(* IEC 61131-3 sources: Lasal-MCP/examples/SampleSource/LASALScreenAdvancedSolution/LASALScreenAdvancedSolution/LASALScreenAdvacnedSolution/Stations/Terminal/HMI/Class/IconDestList, 1 file *)

(* ---- IconDestList.st ---- *)
(*!
<Class
	Name               = "IconDestList"
	Revision           = "0.0"
	RealtimeTask       = "false"
	CyclicTask         = "false"
	BackgroundTask     = "false"
	Sigmatek           = "false"
	OSInterface        = "false"
	HighPriority       = "false"
	Automatic          = "false"
	UpdateMode         = "Prescan"
	SharedCommandTable = "true"
	Objectsize         = "(540,420)">
	<Channels>
		<Client Name="_Grafix" Required="false" Internal="false"/>
		<Client Name="DragDropArea" Required="true" Internal="false"/>
		<Client Name="SigCLib" Required="false" Internal="false"/>
	</Channels>
	<Network Name="IconDestList">
		<!-- List of Components in this network -->
		<Components>
			<Object
				Name       = "_base"
				Class      = "_ScrollArea2"
				Position   = "(218,120)"
				Visualized = "true"
				Remotely   = "true">
				<Channels>
					<Server Name="ActPos"/>
					<Server Name="Refresh"/>
					<Server Name="Server0"/>
					<Client Name="ExtendedScrollBar" Value="0"/>
					<Client Name="LineHighness"/>
					<Client Name="LineWidth"/>
					<Client Name="Lse"/>
					<Client Name="VerticalLevel"/>
				</Channels>
			</Object>
		</Components>
		<Comments>
		</Comments>
		<!-- List of Connections in this network -->
		<Connections>
			<Connection Source="this.Server0" Destination="_base.Server0" Vertices="(886,210),(714,210),"/>
			<Connection Source="this.Refresh" Destination="_base.Refresh" Vertices="(886,270),(714,270),"/>
			<Connection Source="this.ActPos" Destination="_base.ActPos" Vertices="(886,330),(714,330),"/>
			<Connection Source="_base.Lse" Destination="this.Lse" Vertices="(218,210),(38,210),"/>
			<Connection Source="_base.VerticalLevel" Destination="this.VerticalLevel" Vertices="(218,270),(38,270),"/>
			<Connection Source="_base.LineWidth" Destination="this.LineWidth" Vertices="(218,330),(38,330),"/>
		</Connections>
		<!-- Headerfiles -->
		<Options>
		</Options>
	</Network>
</Class>
*)
#pragma using _ScrollArea2

IconDestList : CLASS
: _ScrollArea2
  //Servers:
  //Clients:
	DragDropArea 	: CltChCmd_DragDropArea;
	_Grafix 	: CltChCmd__Grafix;
	SigCLib 	: CltChCmd_SigCLib;
  //Variables:
		TextColor 	: _COLOR;
		FrameColor 	: _COLOR;
		BackgroundColor 	: _COLOR;
		myPioScroll 	: _SCROLL;
		myImageRoom 	: _ROOM;
		Lines : ARRAY [0..100] OF DINT;

		pLSEpio 	: ^_IO;
  //Functions:

	FUNCTION VIRTUAL GLOBAL Init;
				//! <Function Comment="[#ENGLISH]&#13;&#10;method is called cyclic during object is on screen&#13;&#10;&#13;&#10;pio ....... pointer to io information&#13;&#10;input .... TRUE it&apos;s an input / FALSE it&apos;s an output&#13;&#10;" Name="IF_Run"/>
	FUNCTION __CDECL VIRTUAL GLOBAL IF_Run
		VAR_INPUT
			pio 	: ^_IO;			//! <Variable Comment="pointer to _IO information given by LSE" Name="IF_Run.pio"/>
			input 	: BOOL;			//! <Variable Comment="TRUE it&apos;s an input&#13;&#10;FALSE it&apos;s an output" Name="IF_Run.input"/>
		END_VAR;
				//! <Function Comment="method is called every time when redraw of a single line is necessary.&#13;&#10;" Name="Line"/>
	FUNCTION __CDECL VIRTUAL GLOBAL Line
		VAR_INPUT
			ps 	: ^_SCROLL;			//! <Variable Comment="pointer to structure _SCROLL" Name="Line.ps"/>
			pr 	: ^_ROOM;			//! <Variable Comment="pointer to place where line should be drawn" Name="Line.pr"/>
			line 	: UINT;			//! <Variable Comment="16 bit linenumber " Name="Line.line"/>
			state 	: BOOL;			//! <Variable Comment="line is selected (true) or passive (false)" Name="Line.state"/>
		END_VAR;

	FUNCTION GLOBAL GetDimensionDestScroll
		VAR_OUTPUT
			pScroll 	: ^_SCROLL;
		END_VAR;

	FUNCTION GLOBAL InsertIcon
		VAR_INPUT
			IconNo 	: DINT;
			pEvent 	: ^_EVENT;
		END_VAR;
  //Tables:
	FUNCTION @STD
		VAR_OUTPUT
			ret_code	: CONFSTATES;
		END_VAR;
	FUNCTION GLOBAL TAB @CT_;
END_CLASS;

#pragma usingLtd _Grafix
#pragma usingLtd DragDropArea
#pragma usingLtd SigCLib

FUNCTION VIRTUAL GLOBAL IconDestList::Init
VAR
	index : DINT;
END_VAR

  if (_FirstScan = TRUE) then

    for index := 0 to (100) do  // icon 99 from ImageScheme
      Lines[index] := 99;
    end_for;

    pLSEpio := NIL;

    Scroll.position.no := 10; // nummber of Lines
    Scroll.line_height := 75; // height of the line

    TextColor       := _Grafix.MakeColor(backcolor:= INVISIBLE,
                                         frontcolor:= BLACK);

    FrameColor      := _Grafix.MakeColor(backcolor:= INVISIBLE,
                                         frontcolor:= INVISIBLE);

    BackgroundColor := _Grafix.MakeColor(backcolor:= INVISIBLE,
                                         frontcolor:= INVISIBLE);
  end_if;

END_FUNCTION

FUNCTION __CDECL VIRTUAL GLOBAL IconDestList::Line
	VAR_INPUT
		ps 	: ^_SCROLL;
		pr 	: ^_ROOM;
		line 	: UINT;
		state 	: BOOL;
	END_VAR
  VAR
    att       :_ATTRIB;
    schemeNo  : UDINT;
    lineNo    : ARRAY [0..10] of CHAR;
    pImage    : ^_BMP;
  END_VAR

  _memcpy(ptr1:= #myPioScroll, ptr2:= ps, cntr:= sizeof(_SCROLL));

  if (line < Scroll.position.no) then

   ps^.line_height := 75;

   att := T_SOLID or T_COPY or T_PROP or T_LEFTBOUND;

   schemeNo := get_no_by_label(p0:= "DragDrop", x1:= IMAGESCHEME, x2:= 0);

   if (schemeNo = DEFSCOPE) then
     TRACE("Image not found in ImageScheme 'DragDrop'");
     return;
   end_if;

   pImage$^void := NewDoScheme(x0:= IMAGESCHEME,
                               x1:= Lines[line],
                               x2:= schemeNo);

   if (pImage <> NIL) then

     myImageRoom.xy1.x := pr^.xy1.x;
     myImageRoom.xy1.y := pr^.xy1.y;
     myImageRoom.xy2.x := pr^.xy1.x + to_int(Scroll.line_height);
     myImageRoom.xy2.y := pr^.xy2.y;

     out_zoom_BMP(p0:= #myImageRoom,
                  p1:= pImage,
                  x2:= att);

     // insert line no
     myImageRoom.xy1.x := pr^.xy1.x + 76;
     myImageRoom.xy1.y := pr^.xy1.y;
     myImageRoom.xy2.x := pr^.xy1.x + 96;
     myImageRoom.xy2.y := pr^.xy2.y;

     _memset(dest:= #lineNo[0],
             usByte:= 0,
             cntr:= sizeof(lineNo));

     SigCLib.IToA(val:= line,
                  dst:= #lineNo[0],
                  base:= 10);

     if (pLSEpio = NIL) then
       return;
     end_if;

     OutTextAlign(p0:= #lineNo[0],
                  x1:= 0,
                  p1:= #myImageRoom,
                  x2:= pLSEpio^.font,
                  x3:= pLSEpio^.attrib,
                  x9:= pLSEpio^.frametype,
                  x4:= TextColor,
                  x5:= FrameColor,
                  x6:= BackgroundColor,
                  x7:= 1);
   else
     TRACE("Image not found in ImageScheme 'DragDrop'");
   end_if;

  end_if;

END_FUNCTION

FUNCTION GLOBAL IconDestList::GetDimensionDestScroll
	VAR_OUTPUT
		pScroll 	: ^_SCROLL;
	END_VAR

  pScroll := #myPioScroll;

END_FUNCTION

FUNCTION GLOBAL IconDestList::InsertIcon
	VAR_INPUT
		IconNo 	: DINT;
		pEvent 	: ^_EVENT;
	END_VAR
  VAR
  	insertNo : DINT;
  END_VAR

  insertNo := ((pEvent^.dot.y - myPioScroll.out_room.xy1.y)
                / Scroll.line_height) + Scroll.position.begin;

  //Insert in List
  Lines[insertNo] := IconNo;

  LetsDraw := TRUE;

  Refresh := 1;

END_FUNCTION

FUNCTION __CDECL VIRTUAL GLOBAL IconDestList::IF_Run
	VAR_INPUT
		pio 	: ^_IO;
		input 	: BOOL;
	END_VAR

  pLSEpio := pio;
  _ScrollArea2::IF_Run(pio:= pio, input:= input);

END_FUNCTION
